// TIA Portal V17 export
FUNCTION_BLOCK "Sub_FB"   // FB2, LAD
   VAR_INPUT
      Start : Bool;
      Block : Bool;
   END_VAR
   VAR_OUTPUT
      Run : Bool;
   END_VAR
   VAR
      Latch : Bool;
   END_VAR
BEGIN

REGION Network 1
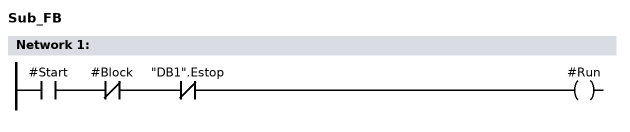
   RUNG wire#powerrail
      Contact( #Start )
      I_Contact( #Block )
      I_Contact( "DB1".Estop )
      Coil( #Run )
   END_RUNG
   // the same network as SCL:
   #Run := #Start AND NOT #Block AND NOT "DB1".Estop;
END_REGION
END_FUNCTION_BLOCK
